// TIA Portal V20 export
VAR_GLOBAL   // PLC tag table "COGNEX_FOLIE_L"
   "COG_FOLIE_L_COG_FOLIE_L_is3800-TriggerEnable" AT %Q5.0 : Bool;
   "COG_FOLIE_L_is3800-Trigger" AT %Q5.1 : Bool;
   "COG_FOLIE_L_is3800-ClearExposureComplete" AT %Q5.2 : Bool;
   "COG_FOLIE_L_is3800-Set Offline" AT %Q5.7 : Bool;
   "COG_FOLIE_L_is3800-TriggerReady" AT %I14.0 : Bool;
   "COG_FOLIE_L_is3800-TriggerAck" AT %I14.1 : Bool;
   "COG_FOLIE_L_is3800-ExposureComplete" AT %I14.2 : Bool;
   "COG_FOLIE_L_is3800-AcquCOG_FOLIE_L_isitionError" AT %I14.3 : Bool;
   "COG_FOLIE_L_is3800-Offline Reason" AT %I14.4 : Bool;
   "COG_FOLIE_L_is3800-Offline Reason(1)" AT %I14.5 : Bool;
   "COG_FOLIE_L_is3800-Offline Reason(2)" AT %I14.6 : Bool;
   "COG_FOLIE_L_is3800-Online" AT %I14.7 : Bool;
   "COG_FOLIE_L_is3800-AcquCOG_FOLIE_L_isitionID" AT %IW16 : Int;
   "COG_FOLIE_L_is3800-BufferResultsEnable" AT %Q6.0 : Bool;
   "COG_FOLIE_L_is3800-InspectionResultsAck" AT %Q6.1 : Bool;
   "COG_FOLIE_L_is3800-SetUserData" AT %Q6.2 : Bool;
   "COG_FOLIE_L_is3800-ExecuteCommand/JobLoad" AT %Q6.3 : Bool;
   "COG_FOLIE_L_is3800-ClearError" AT %Q6.7 : Bool;
   "COG_FOLIE_L_is3800-Reserved" AT %I18.0 : Bool;
   "COG_FOLIE_L_is3800-InspectionCompleted" AT %I18.1 : Bool;
   "COG_FOLIE_L_is3800-ResultsBufferOverrun" AT %I18.2 : Bool;
   "COG_FOLIE_L_is3800-ResultsValid" AT %I18.3 : Bool;
   "COG_FOLIE_L_is3800-CommandExecuting" AT %I18.4 : Bool;
   "COG_FOLIE_L_is3800-CommandCompleted" AT %I18.5 : Bool;
   "COG_FOLIE_L_is3800-CommandFailed" AT %I18.6 : Bool;
   "COG_FOLIE_L_is3800-SetUserDataAck" AT %I18.7 : Bool;
   "COG_FOLIE_L_is3800-ResultsPassed (Job)" AT %I19.0 : Bool;
   "COG_FOLIE_L_is3800-SystemValidated" AT %I19.1 : Bool;
   "COG_FOLIE_L_is3800-Error" AT %I19.7 : Bool;
   "COG_FOLIE_L_is3800-ErrorCode" AT %IW20 : Word;
   "COG_FOLIE_L_is3800-CommandID" AT %QW130 : Word;
   "COG_FOLIE_L_is3800-Current Job ID" AT %IW140 : Word;
   "COG_FOLIE_L_is3800-CommandResultCode" AT %IW142 : Word;
   "COG_FOLIE_L_is3800-ExternalEvent[0]" AT %Q7.0 : Bool;
   "COG_FOLIE_L_is3800-ExternalEvent[1]" AT %Q7.1 : Bool;
   "COG_FOLIE_L_is3800-ExternalEvent[2]" AT %Q7.2 : Bool;
   "COG_FOLIE_L_is3800-ExternalEvent[3]" AT %Q7.3 : Bool;
   "COG_FOLIE_L_is3800-ExternalEvent[4]" AT %Q7.4 : Bool;
   "COG_FOLIE_L_is3800-ExternalEvent[5]" AT %Q7.5 : Bool;
   "COG_FOLIE_L_is3800-ExternalEvent[6]" AT %Q7.6 : Bool;
   "COG_FOLIE_L_is3800-ExternalEvent[7]" AT %Q7.7 : Bool;
   "COG_FOLIE_L_is3800-ExternalEventAck[0]" AT %I7.0 : Bool;
   "COG_FOLIE_L_is3800-ExternalEventAck[1]" AT %I7.1 : Bool;
   "COG_FOLIE_L_is3800-ExternalEventAck[2]" AT %I7.2 : Bool;
   "COG_FOLIE_L_is3800-ExternalEventAck[3]" AT %I7.3 : Bool;
   "COG_FOLIE_L_is3800-ExternalEventAck[4]" AT %I7.4 : Bool;
   "COG_FOLIE_L_is3800-ExternalEventAck[5]" AT %I7.5 : Bool;
   "COG_FOLIE_L_is3800-ExternalEventAck[6]" AT %I7.6 : Bool;
   "COG_FOLIE_L_is3800-ExternalEventAck[7]" AT %I7.7 : Bool;
   "COG_FOLIE_L_is3800-UserData[0]" AT %QB132 : Byte;
   "COG_FOLIE_L_is3800-UserData[1]" AT %QB133 : Byte;
   "COG_FOLIE_L_is3800-UserData[2]" AT %QB134 : Byte;
   "COG_FOLIE_L_is3800-UserData[3]" AT %QB135 : Byte;
   "COG_FOLIE_L_is3800-UserData[4]" AT %QB136 : Byte;
   "COG_FOLIE_L_is3800-UserData[5]" AT %QB137 : Byte;
   "COG_FOLIE_L_is3800-UserData[6]" AT %QB138 : Byte;
   "COG_FOLIE_L_is3800-UserData[7]" AT %QB139 : Byte;
   "COG_FOLIE_L_is3800-UserData[8]" AT %QB140 : Byte;
   "COG_FOLIE_L_is3800-UserData[9]" AT %QB141 : Byte;
   "COG_FOLIE_L_is3800-UserData[10]" AT %QB142 : Byte;
   "COG_FOLIE_L_is3800-UserData[11]" AT %QB143 : Byte;
   "COG_FOLIE_L_is3800-UserData[12]" AT %QB144 : Byte;
   "COG_FOLIE_L_is3800-UserData[13]" AT %QB145 : Byte;
   "COG_FOLIE_L_is3800-UserData[14]" AT %QB146 : Byte;
   "COG_FOLIE_L_is3800-UserData[15]" AT %QB147 : Byte;
   "COG_FOLIE_L_is3800-InspectionID" AT %IW144 : Word;
   "COG_FOLIE_L_is3800-InspectionResultsCode" AT %IW146 : Int;
   "COG_FOLIE_L_is3800-InspectionResults[0]" AT %IB148 : Byte;
   "COG_FOLIE_L_is3800-InspectionResults[1]" AT %IB149 : Byte;
   "COG_FOLIE_L_is3800-InspectionResults[2]" AT %IB150 : Byte;
   "COG_FOLIE_L_is3800-InspectionResults[3]" AT %IB151 : Byte;
   "COG_FOLIE_L_is3800-InspectionResults[4]" AT %IB152 : Byte;
   "COG_FOLIE_L_is3800-InspectionResults[5]" AT %IB153 : Byte;
   "COG_FOLIE_L_is3800-InspectionResults[6]" AT %IB154 : Byte;
   "COG_FOLIE_L_is3800-InspectionResults[7]" AT %IB155 : Byte;
   "COG_FOLIE_L_is3800-InspectionResults[8]" AT %IB156 : Byte;
   "COG_FOLIE_L_is3800-InspectionResults[9]" AT %IB157 : Byte;
   "COG_FOLIE_L_is3800-InspectionResults[10]" AT %IB158 : Byte;
   "COG_FOLIE_L_is3800-InspectionResults[11]" AT %IB159 : Byte;
   "COG_FOLIE_L_is3800-InspectionResults[12]" AT %IB160 : Byte;
   "COG_FOLIE_L_is3800-InspectionResults[13]" AT %IB161 : Byte;
   "COG_FOLIE_L_is3800-InspectionResults[14]" AT %IB162 : Byte;
   "COG_FOLIE_L_is3800-InspectionResults[15]" AT %IB163 : Byte;
END_VAR
